// TIA Portal V19 export
FUNCTION_BLOCK "SCALING"   // FB3, FBD
{ S7_Optimized_Access := 'TRUE' }
// stored: MemoryReserve 100, SetENOAutomatically false
   VAR_INPUT
      RAW_MIN : Int;
      RAW_MAX : Int;
      INPUT : Int;
      SCALE_MIN : Real;
      SCALE_MAX : Real;
   END_VAR
   VAR_OUTPUT
      SCALE_OUT : Real;
   END_VAR
   VAR
      TEMP : Real;
   END_VAR
BEGIN

REGION Network 1
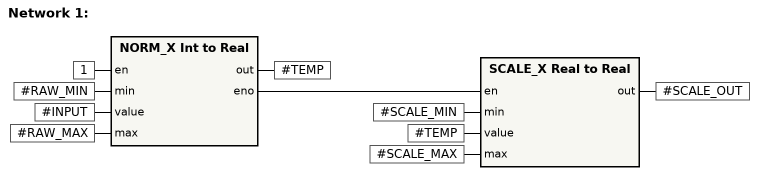
   IF 1 THEN
       #TEMP := NORM_X(MIN := #RAW_MIN, VALUE := #INPUT, MAX := #RAW_MAX);
       #SCALE_OUT := SCALE_X(MIN := #SCALE_MIN, VALUE := #TEMP, MAX := #SCALE_MAX);
   END_IF;
END_REGION
END_FUNCTION_BLOCK
